(* IEC 61131-3 sources: model-first-plc-agent-ai/results/T2-W-08, 2 files *)

(* ---- a1_code.st ---- *)
FUNCTION_BLOCK FillingRuntime
VAR_INPUT
    start : BOOL;
    stop : BOOL;
    LSH : BOOL;
    LSHH : BOOL;
    TimerDuration : TIME;
END_VAR
VAR_OUTPUT
    fill_valve : BOOL;
    discharge_valve : BOOL;
END_VAR
VAR
    x0 : BOOL := TRUE;
    x1 : BOOL := FALSE;
    t1 : BOOL;
    t2 : BOOL;
    timer_done : BOOL := FALSE;
    FillingTimer : TON;
END_VAR

(* Evaluate the start transition from the current situation. *)
t1 := x0 AND start AND NOT stop AND NOT LSHH;

(* Start timing in the scan that activates x1. *)
FillingTimer(
    IN := x1 OR t1,
    PT := TimerDuration
);

(* The owned condition is FALSE at activation of x1. *)
timer_done := x1 AND FillingTimer.Q;

(* Evaluate the return transition before changing the situation. *)
t2 := x1 AND (stop OR LSHH OR timer_done);

IF t2 THEN
    x0 := TRUE;
    x1 := FALSE;
ELSIF t1 THEN
    x0 := FALSE;
    x1 := TRUE;
END_IF;

(* Reset the nonretentive timer when its owning step is inactive. *)
IF NOT x1 THEN
    FillingTimer(IN := FALSE, PT := TimerDuration);
    timer_done := FALSE;
END_IF;

fill_valve := x1;
discharge_valve := FALSE;

END_FUNCTION_BLOCK

PROGRAM Main
VAR
    StartCommand AT %IX100.0 : BOOL;
    StopCommand AT %IX100.1 : BOOL;
    LSH AT %IX100.2 : BOOL;
    LSHH AT %IX100.3 : BOOL;
    FillValve AT %QX100.0 : BOOL;
    DischargeValve AT %QX100.1 : BOOL;
END_VAR
VAR
    (* Configurable filling interval. *)
    TimerDuration : TIME := T#10s;
    StartEdge : R_TRIG;
    FillingControl : FillingRuntime;
END_VAR

StartEdge(CLK := StartCommand);

FillingControl(
    start := StartEdge.Q,
    stop := StopCommand,
    LSH := LSH,
    LSHH := LSHH,
    TimerDuration := TimerDuration
);

FillValve := FillingControl.fill_valve;
DischargeValve := FillingControl.discharge_valve;

END_PROGRAM

(* ---- a2_code.st ---- *)
FUNCTION_BLOCK FB_TimedFilling
VAR_INPUT
    StartCommand : BOOL;
    StopCommand : BOOL;
    LSH : BOOL;
    LSHH : BOOL;
    TimerDuration : TIME;
END_VAR
VAR_OUTPUT
    fill_valve : BOOL;
    discharge_valve : BOOL;
END_VAR
VAR
    StartEdge : R_TRIG;
    FillingTimer : TON;
    ActiveState : INT := 0;
    start : BOOL;
    stop : BOOL;
    timer_done : BOOL := FALSE;
END_VAR

StartEdge(CLK := StartCommand);
start := StartEdge.Q;
stop := StopCommand;

IF stop THEN
    ActiveState := 0;
ELSE
    CASE ActiveState OF
        0:
            IF start THEN
                ActiveState := 1;
            END_IF;
        1:
            ActiveState := 1;
    ELSE
        ActiveState := 0;
    END_CASE;
END_IF;

FillingTimer(
    IN := (ActiveState = 1),
    PT := TimerDuration
);
timer_done := FillingTimer.Q;

IF ActiveState = 1 THEN
    IF stop OR timer_done OR LSHH THEN
        ActiveState := 0;
        FillingTimer(IN := FALSE, PT := TimerDuration);
        timer_done := FALSE;
    END_IF;
END_IF;

fill_valve := (ActiveState = 1);
discharge_valve := FALSE;

END_FUNCTION_BLOCK

PROGRAM Main
VAR
    StartCommand AT %IX100.0 : BOOL;
    StopCommand AT %IX100.1 : BOOL;
    LSH AT %IX100.2 : BOOL;
    LSHH AT %IX100.3 : BOOL;
    FillValve AT %QX100.0 : BOOL;
    DischargeValve AT %QX100.1 : BOOL;
END_VAR
VAR
    FillingControl : FB_TimedFilling;
    TimerDuration : TIME := T#10s;
END_VAR

FillingControl(
    StartCommand := StartCommand,
    StopCommand := StopCommand,
    LSH := LSH,
    LSHH := LSHH,
    TimerDuration := TimerDuration
);

FillValve := FillingControl.fill_valve;
DischargeValve := FillingControl.discharge_valve;

END_PROGRAM
